// Halbzeugdaten des aktiven Programms.
{attribute 'pack_mode' := '1'}
TYPE ST_Material :
STRUCT
    fDiameter_mm : LREAL;
    fWall_mm : LREAL; // 0 = Vollmaterial
    fYield_MPa : LREAL; // Rp0,2
    fForceLimit_N : LREAL;
END_STRUCT
END_TYPE

(* stored: Version 1.1.0.1
   DUT ST_Material: Id {1946f580-3cae-445c-9069-80ba1f71f6fa} *)
